(* IEC 61131-3 sources: guidance-for-physical-ai-production-designer-on-aws/source/plan2cell/examples/cell_2robot/plc/codesys/head/DUT, 8 files *)

(* ---- E_CellError.st ---- *)
(*
 * E_CellError
 *
 * Fault codes of the cell (FB_Cell.eError), the robot drivers (FB_VassRobot.eError)
 * and the zone arbiter (FB_ZoneArbiter.eFault). ERR_NONE = no fault.
 *)

TYPE E_CellError :
(
    ERR_NONE                := 0,

    (* VASS bring-up and job handshake (FB_VassRobot) *)
    ERR_SAFETY_TIMEOUT      := 10,      (* SafeIn0.0 / SafeIn1.4 not reported *)
    ERR_DRIVES_TIMEOUT      := 11,      (* DrivesOn not reported *)
    ERR_EXT_TIMEOUT         := 12,      (* EXT mode not reported *)
    ERR_NOT_READY           := 13,      (* robot not Ready (or JobAck stuck) before a job *)
    ERR_ACK_TIMEOUT         := 14,      (* no JobAck after JobRequest *)
    ERR_ECHO_MISMATCH       := 15,      (* echoed job number <> requested job number *)
    ERR_START_TIMEOUT       := 16,      (* ProgRunning not reported after ProgStart *)
    ERR_ROBOT_STOPPED       := 17,      (* ProgRunning dropped without ProgFinished (T_STOP_DEBOUNCE) *)
    ERR_ROBOT_ERROR         := 18,      (* robot reports Error *)
    ERR_SAFETY_LOST         := 19,      (* safe status lost while up *)
    ERR_STOP_TIMEOUT        := 20,      (* robot still running after Stop + Cancel *)
    ERR_RESET_FAILED        := 21,      (* robot still in error after Reset *)
    ERR_DRIVES_LOST         := 22,      (* DrivesOn lost while up *)
    ERR_UNEXPECTED_RUN      := 23,      (* ProgRunning reported outside a job (off / bring-up / idle) *)

    (* zone protocol and supervision (FB_ZoneArbiter, FB_Cell) *)
    ERR_OP_WATCHDOG         := 30,      (* op took longer than aOps[].tLimit *)
    ERR_ZONE_WAIT_TIMEOUT   := 31,      (* zone wait past aOps[].tZoneDeadline since cycle start *)
    ERR_STEP_SEQUENCE       := 32,      (* op index did not advance by exactly +1, or 0 between two ops *)
    ERR_REQ_MISMATCH        := 33,      (* REQUEST <> mask of the reported op (debounced) *)
    ERR_TICKET_SKIPPED      := 34,      (* own ticket for another op, or zone consumed (debounced) *)
    ERR_PROGRAM_INCOMPLETE  := 35,      (* job done but last op index <> op count *)
    ERR_RELEASE_INVALID     := 36,      (* REQUEST dropped by a robot that is not running OK *)
    ERR_ROBOT_STALLED       := 37,      (* zone op without REQUEST and grant, or op index 0 too long *)
    ERR_UNEXPECTED_REQUEST  := 38,      (* holder raised bits it was not granted *)
    ERR_TICKETS_LEFT        := 39,      (* cycle done with unconsumed tickets *)
    ERR_HOME_FAILED         := 40,      (* blind homing did not reach the home pose *)
    ERR_HANDSHAKE           := 41,      (* op index changed while a grant was held (4-phase violated) *)
    ERR_ZONE_BYPASSED       := 42,      (* zone / permit op left without ever being granted *)

    (* operator *)
    ERR_OPERATOR_STOP       := 50       (* bStop *)
);
END_TYPE

(* ---- E_CellState.st ---- *)
(*
 * E_CellState
 *
 * States of the cell controller FB_Cell.
 *)

TYPE E_CellState :
(
    CS_INIT                 := 0,       (* robots off *)
    CS_BRINGUP              := 10,      (* all robots: SAFETY_ENABLE -> DRIVES_ON -> MODE_EXT -> IDLE *)
    CS_HOMING_SELECT        := 20,      (* pick robot(s) not at home *)
    CS_HOMING_RUN           := 21,      (* blind homing with HOME_FOLGE *)
    CS_READY                := 30,      (* all robots at home, waiting for start / auto-run *)
    CS_START_JOBS           := 40,      (* production Folge commanded on every active robot *)
    CS_RUNNING              := 50,      (* robots run autonomously, zones arbitrated *)
    CS_CYCLE_DONE           := 60,      (* pause T_CYCLE_PAUSE before the next cycle *)
    CS_ABORTING             := 80,      (* grants dropped, Stop + Cancel to every busy robot *)
    CS_RECOVERY             := 85,      (* after an abort mid-cycle, or a start-up with an active robot
                                           away from home: wait for bRecoveryConfirm *)
    CS_RESETTING            := 90,      (* Reset to robots in error (an operator stop cancels it) *)
    CS_ERROR                := 99       (* latched until bReset *)
);
END_TYPE

(* ---- E_GrantPolicy.st ---- *)
(*
 * E_GrantPolicy
 *
 * Zone grant policy of FB_ZoneArbiter (GVL_Cell.GRANT_POLICY).
 *)

TYPE E_GrantPolicy :
(
    GP_PLANNED  := 0,       (* zone granted only to its next ticket holder (BT order) *)
    GP_FCFS     := 1        (* oldest request first - BT order NOT enforced *)
);
END_TYPE

(* ---- E_RobotState.st ---- *)
(*
 * E_RobotState
 *
 * States of the VASS driver FB_VassRobot (one robot).
 *)

TYPE E_RobotState :
(
    RS_OFF                  := 0,       (* outputs off, waiting for bPowerOn *)
    RS_SAFETY_ENABLE        := 1,       (* SafeOut0/1 set, waiting for safe status *)
    RS_DRIVES_ON            := 2,       (* DrivesOn requested *)
    RS_MODE_EXT             := 3,       (* EXT mode requested *)
    RS_IDLE                 := 10,      (* up, no job *)
    RS_JOB_WAIT_READY       := 20,      (* waiting for Ready and no JobAck *)
    RS_JOB_SEND             := 21,      (* job number + JobRequest, waiting for JobAck *)
    RS_JOB_START            := 22,      (* ProgStart pulse *)
    RS_JOB_WAIT_RUNNING     := 23,      (* waiting for ProgRunning (or ProgFinished) *)
    RS_JOB_RUNNING          := 24,      (* program running *)
    RS_JOB_DONE             := 25,      (* ProgFinished seen, bJobDone set *)
    RS_STOPPING             := 30,      (* Stop + Cancel held *)
    RS_RESET                := 40,      (* Reset held *)
    RS_ERROR                := 99       (* latched until bCmdReset *)
);
END_TYPE

(* ---- ST_OpInfo.st ---- *)
(*
 * ST_OpInfo
 *
 * One op of one robot (GVL_Cell.aOps). Op k of robot r is
 * GVL_Cell.aOps[GVL_Cell.anRobotFirstOp[r] + k - 1].
 *)

TYPE ST_OpInfo :
STRUCT
    nRobot              : INT;      (* robot index, 1-based *)
    nOp                 : INT;      (* op index of that robot, 1-based *)
    dwZoneMask          : DWORD;    (* REQUEST/GRANT mask: zone bits 0..30, bit 31 = permit *)
    nPredFirst          : INT;      (* permit preds: GVL_Cell.aPreds[nPredFirst .. nPredFirst + nPredCount - 1] *)
    nPredCount          : INT;      (* 0 = no permit predecessors *)
    tExpected           : TIME;     (* nominal duration *)
    tLimit              : TIME;     (* op watchdog (from the grant, or from the step change if mask = 0) *)
    tZoneDeadline       : TIME;     (* latest grant time since cycle start *)
    sName               : STRING(32);
END_STRUCT
END_TYPE

(* ---- ST_RobotIn.st ---- *)
(*
 * ST_RobotIn
 *
 * Copy of one robot's input image (robot -> PLC), filled by PLC_PRG from
 * GVL_IO.bySafeIn0_<tag>..bySafeIn7_<tag> and GVL_IO.aVassInputData_<tag>.
 *)

TYPE ST_RobotIn :
STRUCT
    abySafeIn           : ARRAY[0..7] OF BYTE;      (* PROFIsafe FDIO64 safe status *)
    aVassIn             : ARRAY[0..31] OF BYTE;     (* VASS DIO256 status telegram *)
END_STRUCT
END_TYPE

(* ---- ST_RobotOut.st ---- *)
(*
 * ST_RobotOut
 *
 * One robot's output image (PLC -> robot), copied by PLC_PRG to
 * GVL_IO.bySafeOut0_<tag>..bySafeOut7_<tag> and GVL_IO.aVassOutputData_<tag>.
 *)

TYPE ST_RobotOut :
STRUCT
    abySafeOut          : ARRAY[0..7] OF BYTE;      (* PROFIsafe FDIO64 safe commands *)
    aVassOut            : ARRAY[0..31] OF BYTE;     (* VASS DIO256 command telegram *)
END_STRUCT
END_TYPE

(* ---- ST_Ticket.st ---- *)
(*
 * ST_Ticket
 *
 * One (robot, op) reference: a zone ticket in GVL_Cell.aTickets or a permit
 * predecessor in GVL_Cell.aPreds. Both indices are 1-based; 0 = none (dummy row).
 *)

TYPE ST_Ticket :
STRUCT
    nRobot              : INT;      (* robot index 1..GVL_Cell.N_ROBOTS *)
    nOp                 : INT;      (* op index of that robot 1..anRobotOpCount[nRobot] *)
END_STRUCT
END_TYPE
